(* Schneider Machine Expert - Basic project Traffic_light, file version 2.9.0.0 *)
(* ProjectInformations: Name=New project *)

HARDWARE
  Cpu 0: TM221M16R/G
  EthernetConfiguration: NetworkName=M221, IpAllocationMode=FixedAddress, IpAddress=0.0.0.0, SubnetMask=0.0.0.0
  SerialLineConfiguration: Baud=Baud19200, Parity=ParityEven, DataBits=DataBits8, StopBits=StopBits1, PhysicalMedium=PhysicalMediumRs485, TransmissionMode=TransmissionModeModbusRtu, SlaveId=1, Addressing=SlaveAddressing
  MastTask: UsePeriodScanMode=false, PeriodScan=100
  FastTask: Period=255
  CpuBehavior: StartingMode=StartAsPreviousState, AutoSaveRamOnEeprom=true, WatchdogPeriod=250

SYMBOLS  (address, symbol, comment, settings)
  %M1       RED_ONLY_SET
  %M2       RED_PLUS_YELOW_SET
  %M3       GREEN_ONLY_SET
  %M4       GREEN_BLINK_SWITCH
  %M5       GREEN_BLINK_SIG_GEN
  %M6       GREEN_BLINK_SET
  %M7       YELOW_ONLEY_SET
  %M8       DELEY_GREEN_ONLY_SET
  %TM0      RED_UELOW_TON  [Preset=3, Base=OneSecond]
  %TM1      GREEN_TON  [Preset=3, Base=OneSecond]
  %TM2      BLINK_GREAN_TON  [Preset=3, Base=OneSecond]
  %TM3      GREEN_BLINK_SIGNAL_TON  [Preset=1, Base=OneSecond]
  %TM4      GREEN_BLINK_SIGNAL_TOF  [Type=TOF, Preset=1, Base=OneSecond]
  %TM5      RED_ONLEY_ON  [Preset=3, Base=OneSecond]
  %TM6      RED_DELEY  [Preset=1, Base=OneSecond]
  %TM7        [Preset=2, Base=OneSecond]
  %TM8      DELAY_SWITCH_TO_GREEN_ONLEY  [Preset=1, Base=OneSecond]
  %C0         [Preset=3]
  %Q0.0     RED_OUT
  %Q0.1     YELOW_OUT
  %Q0.2     GREEN_OUT

POU New POU
  (* SectionNumber=1 *)

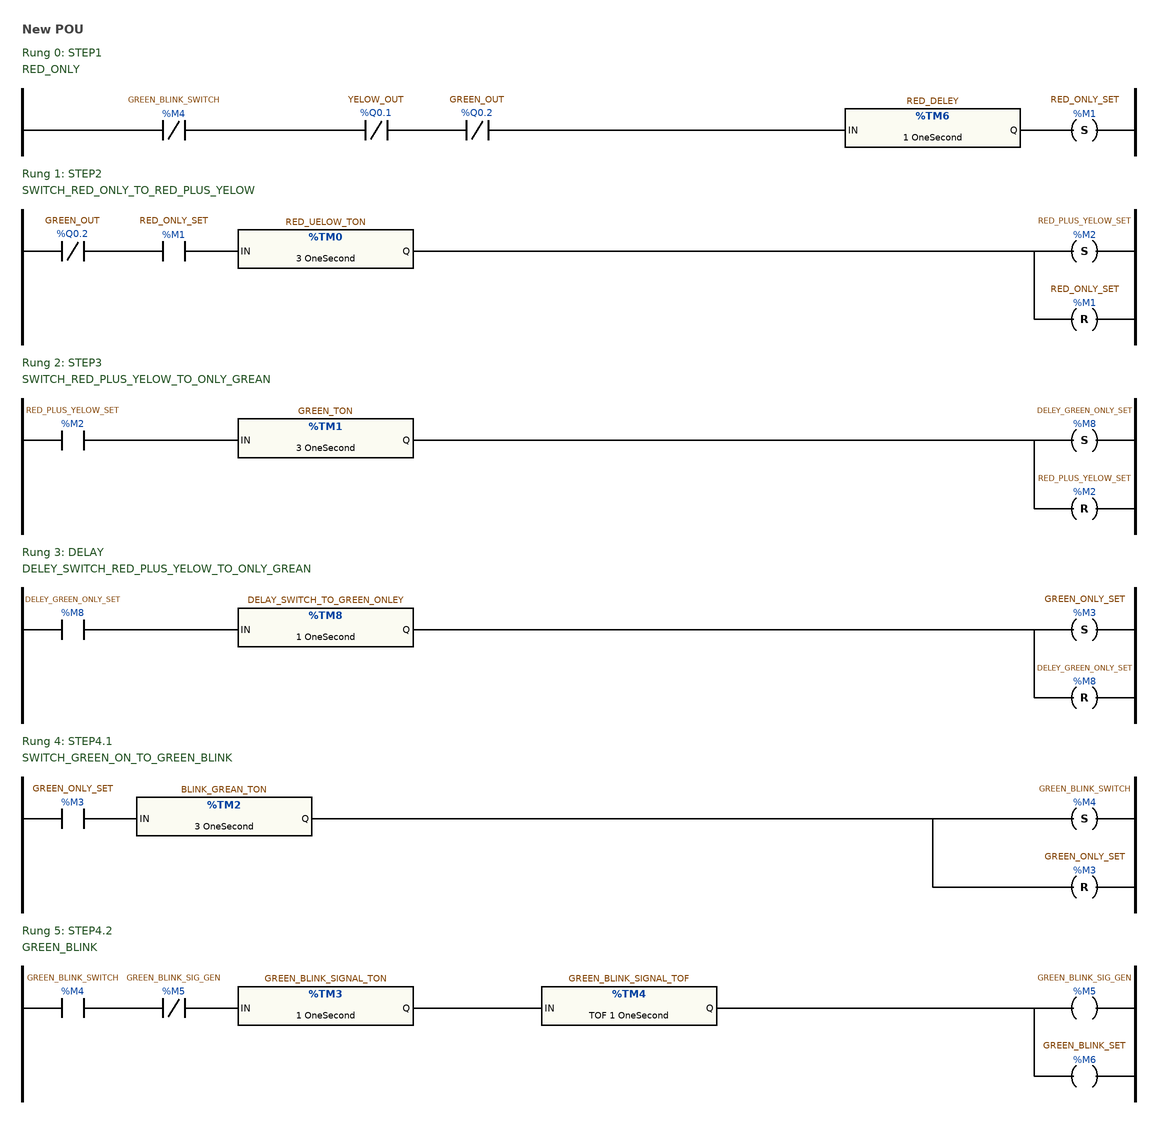

// Rung 0: STEP1
// RED_ONLY
  BLK %TM6                (* RED_DELEY *)
  LDN %M4                 (* GREEN_BLINK_SWITCH *)
  ANDN %Q0.1              (* YELOW_OUT *)
  ANDN %Q0.2              (* GREEN_OUT *)
  IN
  OUT_BLK
  LD Q
  S %M1                   (* RED_ONLY_SET *)
  END_BLK
  // as ST:
  //   RED_DELEY(IN := NOT GREEN_BLINK_SWITCH AND NOT YELOW_OUT AND NOT GREEN_OUT);
  //   IF RED_DELEY.Q THEN RED_ONLY_SET := TRUE; END_IF;

// Rung 1: STEP2
// SWITCH_RED_ONLY_TO_RED_PLUS_YELOW
  BLK %TM0                (* RED_UELOW_TON *)
  LDN %Q0.2               (* GREEN_OUT *)
  AND %M1                 (* RED_ONLY_SET *)
  IN
  OUT_BLK
  LD Q
  S %M2                   (* RED_PLUS_YELOW_SET *)
  R %M1                   (* RED_ONLY_SET *)
  END_BLK
  // as ST:
  //   RED_UELOW_TON(IN := NOT GREEN_OUT AND RED_ONLY_SET);
  //   IF RED_UELOW_TON.Q THEN RED_PLUS_YELOW_SET := TRUE; END_IF;
  //   IF RED_UELOW_TON.Q THEN RED_ONLY_SET := FALSE; END_IF;

// Rung 2: STEP3
// SWITCH_RED_PLUS_YELOW_TO_ONLY_GREAN
  BLK %TM1                (* GREEN_TON *)
  LD %M2                  (* RED_PLUS_YELOW_SET *)
  IN
  OUT_BLK
  LD Q
  S %M8                   (* DELEY_GREEN_ONLY_SET *)
  R %M2                   (* RED_PLUS_YELOW_SET *)
  END_BLK
  // as ST:
  //   GREEN_TON(IN := RED_PLUS_YELOW_SET);
  //   IF GREEN_TON.Q THEN DELEY_GREEN_ONLY_SET := TRUE; END_IF;
  //   IF GREEN_TON.Q THEN RED_PLUS_YELOW_SET := FALSE; END_IF;

// Rung 3: DELAY
// DELEY_SWITCH_RED_PLUS_YELOW_TO_ONLY_GREAN
  BLK %TM8                (* DELAY_SWITCH_TO_GREEN_ONLEY *)
  LD %M8                  (* DELEY_GREEN_ONLY_SET *)
  IN
  OUT_BLK
  LD Q
  S %M3                   (* GREEN_ONLY_SET *)
  R %M8                   (* DELEY_GREEN_ONLY_SET *)
  END_BLK
  // as ST:
  //   DELAY_SWITCH_TO_GREEN_ONLEY(IN := DELEY_GREEN_ONLY_SET);
  //   IF DELAY_SWITCH_TO_GREEN_ONLEY.Q THEN GREEN_ONLY_SET := TRUE; END_IF;
  //   IF DELAY_SWITCH_TO_GREEN_ONLEY.Q THEN DELEY_GREEN_ONLY_SET := FALSE; END_IF;

// Rung 4: STEP4.1
// SWITCH_GREEN_ON_TO_GREEN_BLINK
  BLK %TM2                (* BLINK_GREAN_TON *)
  LD %M3                  (* GREEN_ONLY_SET *)
  IN
  OUT_BLK
  LD Q
  S %M4                   (* GREEN_BLINK_SWITCH *)
  R %M3                   (* GREEN_ONLY_SET *)
  END_BLK
  // as ST:
  //   BLINK_GREAN_TON(IN := GREEN_ONLY_SET);
  //   IF BLINK_GREAN_TON.Q THEN GREEN_BLINK_SWITCH := TRUE; END_IF;
  //   IF BLINK_GREAN_TON.Q THEN GREEN_ONLY_SET := FALSE; END_IF;

// Rung 5: STEP4.2
// GREEN_BLINK
  LD 1
  MULTIFB
  BLK %TM3                (* GREEN_BLINK_SIGNAL_TON *)
  LD 1
  AND %M4                 (* GREEN_BLINK_SWITCH *)
  ANDN %M5                (* GREEN_BLINK_SIG_GEN *)
  IN
  OUT_BLK
  LD Q
  ST %MW2009:X0
  END_BLK
  BLK %TM4                (* GREEN_BLINK_SIGNAL_TOF *)
  LD %MW2009:X0
  IN
  OUT_BLK
  LD Q
  ST %M5                  (* GREEN_BLINK_SIG_GEN *)
  ST %M6                  (* GREEN_BLINK_SET *)
  END_BLK
  MULTIFB
  // as ST:
  //   GREEN_BLINK_SIGNAL_TON(IN := GREEN_BLINK_SWITCH AND NOT GREEN_BLINK_SIG_GEN);
  //   GREEN_BLINK_SIGNAL_TOF(IN := GREEN_BLINK_SIGNAL_TON.Q);
  //   GREEN_BLINK_SIG_GEN := GREEN_BLINK_SIGNAL_TOF.Q;
  //   GREEN_BLINK_SET := GREEN_BLINK_SIGNAL_TOF.Q;

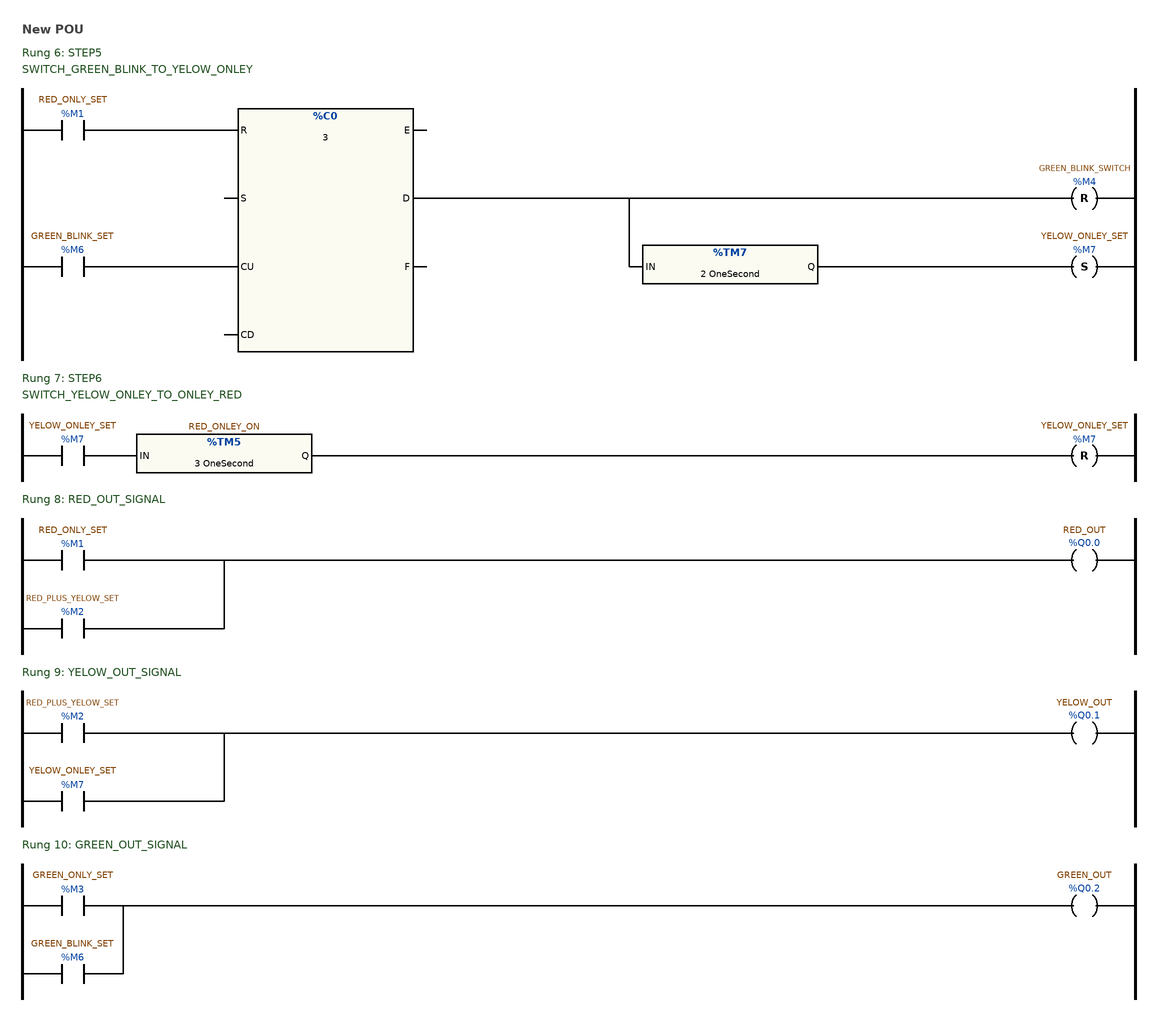

// Rung 6: STEP5
// SWITCH_GREEN_BLINK_TO_YELOW_ONLEY
  LD 1
  MULTIFB
  BLK %C0
  LD 1
  AND %M1                 (* RED_ONLY_SET *)
  R
  LD 1
  AND %M6                 (* GREEN_BLINK_SET *)
  CU
  OUT_BLK
  LD D
  ST %MW2009:X0
  END_BLK
  LD %MW2009:X0
  R %M4                   (* GREEN_BLINK_SWITCH *)
  BLK %TM7
  LD %MW2009:X0
  IN
  OUT_BLK
  LD Q
  S %M7                   (* YELOW_ONLEY_SET *)
  END_BLK
  MULTIFB
  // as ST:
  //   %C0(R := RED_ONLY_SET, CU := GREEN_BLINK_SET);
  //   IF %C0.D THEN GREEN_BLINK_SWITCH := FALSE; END_IF;
  //   %TM7(IN := %C0.D);
  //   IF %TM7.Q THEN YELOW_ONLEY_SET := TRUE; END_IF;

// Rung 7: STEP6
// SWITCH_YELOW_ONLEY_TO_ONLEY_RED
  BLK %TM5                (* RED_ONLEY_ON *)
  LD %M7                  (* YELOW_ONLEY_SET *)
  IN
  OUT_BLK
  LD Q
  R %M7                   (* YELOW_ONLEY_SET *)
  END_BLK
  // as ST:
  //   RED_ONLEY_ON(IN := YELOW_ONLEY_SET);
  //   IF RED_ONLEY_ON.Q THEN YELOW_ONLEY_SET := FALSE; END_IF;

// Rung 8: RED_OUT_SIGNAL
  LD %M1                  (* RED_ONLY_SET *)
  OR %M2                  (* RED_PLUS_YELOW_SET *)
  ST %Q0.0                (* RED_OUT *)
  // as ST:
  //   RED_OUT := RED_ONLY_SET OR RED_PLUS_YELOW_SET;

// Rung 9: YELOW_OUT_SIGNAL
  LD %M2                  (* RED_PLUS_YELOW_SET *)
  OR %M7                  (* YELOW_ONLEY_SET *)
  ST %Q0.1                (* YELOW_OUT *)
  // as ST:
  //   YELOW_OUT := RED_PLUS_YELOW_SET OR YELOW_ONLEY_SET;

// Rung 10: GREEN_OUT_SIGNAL
  LD %M3                  (* GREEN_ONLY_SET *)
  OR %M6                  (* GREEN_BLINK_SET *)
  ST %Q0.2                (* GREEN_OUT *)
  // as ST:
  //   GREEN_OUT := GREEN_ONLY_SET OR GREEN_BLINK_SET;
